Fanuc KAREL source: kt00992.KL

PROGRAM KT00992
%STACKSIZE=65535
%PRIORITY=65535
%NOLOCKGROUP
VAR
P1 : XYZWPR
P2 : XYZWPR
X : REAL
Y : REAL
Z : REAL
W : REAL
P : REAL
R : REAL
-- UNRESOLVED DECLARATIONS (source type spelling not recovered)
-- CFG : TYPE_0x001C (type_u16=0x001C)
BEGIN
P1.X=1.0
P2.Y=2.0
P1.X=1.0
P2.Y=2.0
-- UNRESOLVED_PC line 18 opcodes [27 22 1C 22 22 22 22 22 22 22 76] marker_code=80
END KT00992
